TYPE ST_StationEvents :
STRUCT
	aEvents								: ARRAY [0..100] OF ST_EVENT;	
	
	bFault								: BOOL;
	bCycleStopRequest					: BOOL;
END_STRUCT
END_TYPE

(* stored: Version 1.1.0.1
   DUT ST_StationEvents: Id {496c8842-fa64-4dcc-a4c4-8f89c92f4800} *)
